(* Logix 5000 project; controller CIP_14485201 vendor 1 type 14 code 216 rev 38.11; software revision 38.01; part 5 of 12 *)
(* tags used below, declared in another part *)
   Alarm_Ack : INT[8];   // ALARMS ACKNOWLEDGE BITS
   Alarm_Present : INT[8];   // ALARM MSGS 1-127 PRESENT BITS
   Alarm_Timer : TIMER[128];   // ALARM MSGS 1-127 DELAY TIMERS
(* MainProgram, continued *)

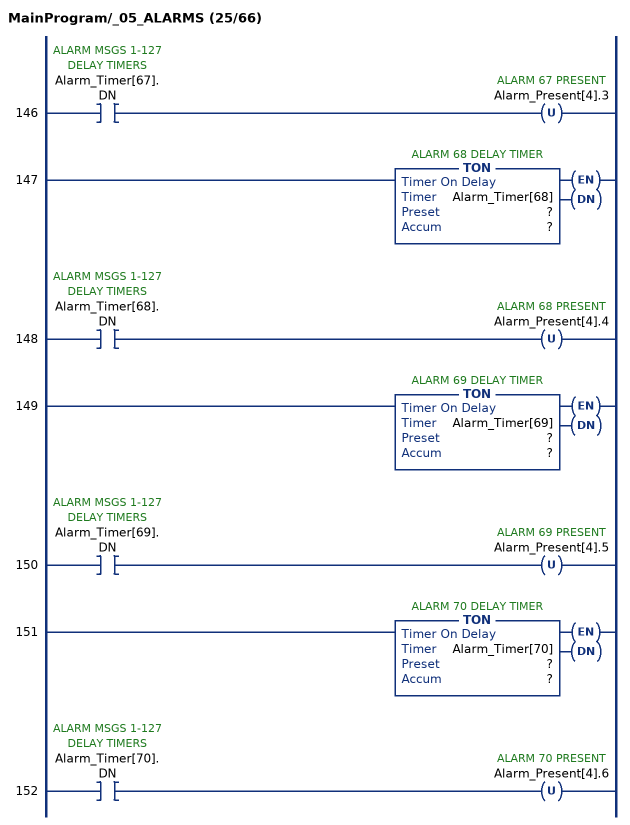
   [picture p52: MainProgram/_05_ALARMS rungs 146-152]
   146: XIC(Alarm_Timer[67].DN)OTU(Alarm_Present[4].3);
   147: TON(Alarm_Timer[68],?,?);
   148: XIC(Alarm_Timer[68].DN)OTU(Alarm_Present[4].4);
   149: TON(Alarm_Timer[69],?,?);
   150: XIC(Alarm_Timer[69].DN)OTU(Alarm_Present[4].5);
   151: TON(Alarm_Timer[70],?,?);
   152: XIC(Alarm_Timer[70].DN)OTU(Alarm_Present[4].6);
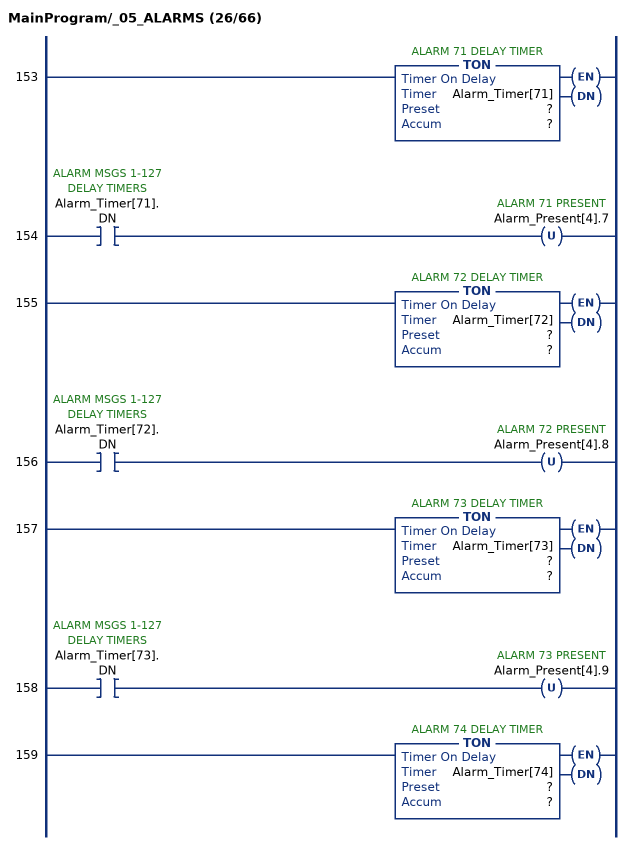
   153: TON(Alarm_Timer[71],?,?);
   154: XIC(Alarm_Timer[71].DN)OTU(Alarm_Present[4].7);
   155: TON(Alarm_Timer[72],?,?);
   156: XIC(Alarm_Timer[72].DN)OTU(Alarm_Present[4].8);
   157: TON(Alarm_Timer[73],?,?);
   158: XIC(Alarm_Timer[73].DN)OTU(Alarm_Present[4].9);
   159: TON(Alarm_Timer[74],?,?);
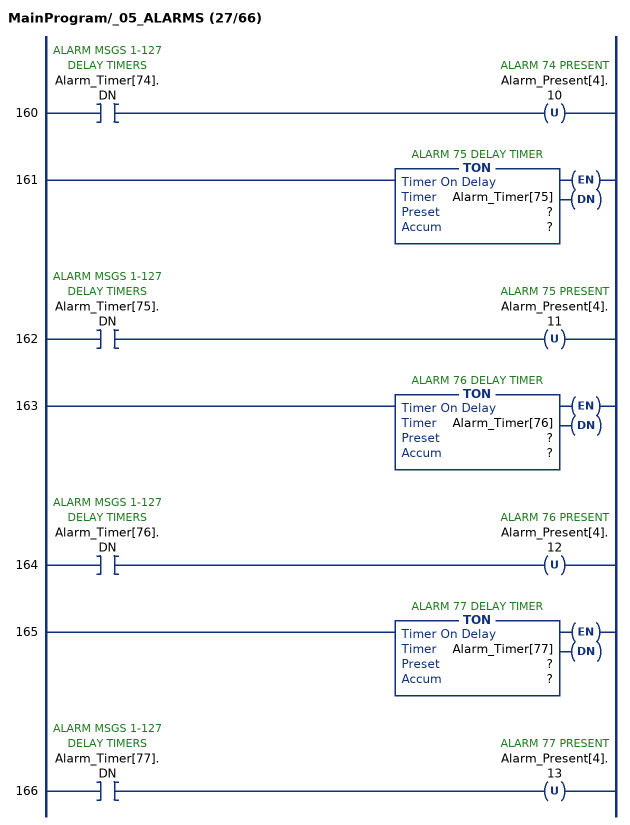
   160: XIC(Alarm_Timer[74].DN)OTU(Alarm_Present[4].10);
   161: TON(Alarm_Timer[75],?,?);
   162: XIC(Alarm_Timer[75].DN)OTU(Alarm_Present[4].11);
   163: TON(Alarm_Timer[76],?,?);
   164: XIC(Alarm_Timer[76].DN)OTU(Alarm_Present[4].12);
   165: TON(Alarm_Timer[77],?,?);
   166: XIC(Alarm_Timer[77].DN)OTU(Alarm_Present[4].13);
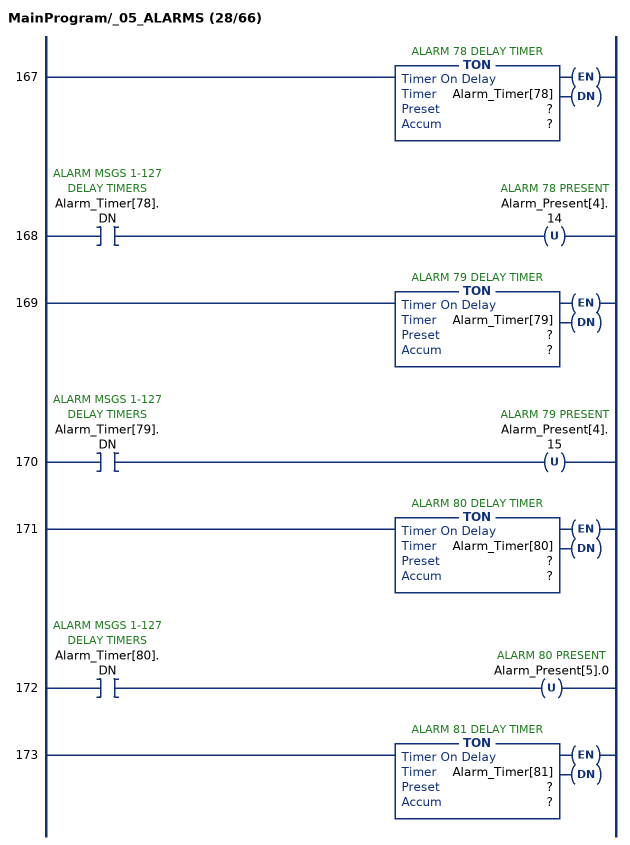
   167: TON(Alarm_Timer[78],?,?);
   168: XIC(Alarm_Timer[78].DN)OTU(Alarm_Present[4].14);
   169: TON(Alarm_Timer[79],?,?);
   170: XIC(Alarm_Timer[79].DN)OTU(Alarm_Present[4].15);
   171: TON(Alarm_Timer[80],?,?);
   172: XIC(Alarm_Timer[80].DN)OTU(Alarm_Present[5].0);
   173: TON(Alarm_Timer[81],?,?);
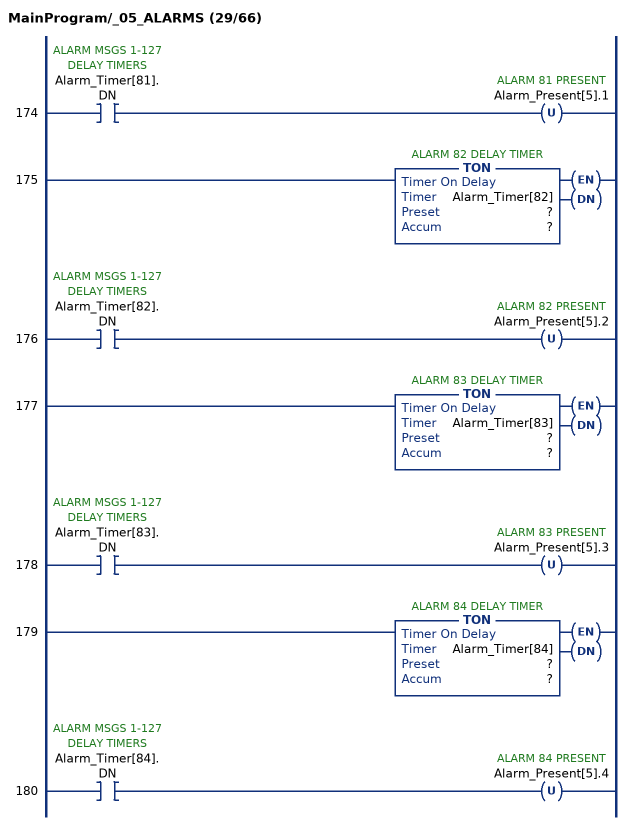
   174: XIC(Alarm_Timer[81].DN)OTU(Alarm_Present[5].1);
   175: TON(Alarm_Timer[82],?,?);
   176: XIC(Alarm_Timer[82].DN)OTU(Alarm_Present[5].2);
   177: TON(Alarm_Timer[83],?,?);
   178: XIC(Alarm_Timer[83].DN)OTU(Alarm_Present[5].3);
   179: TON(Alarm_Timer[84],?,?);
   180: XIC(Alarm_Timer[84].DN)OTU(Alarm_Present[5].4);
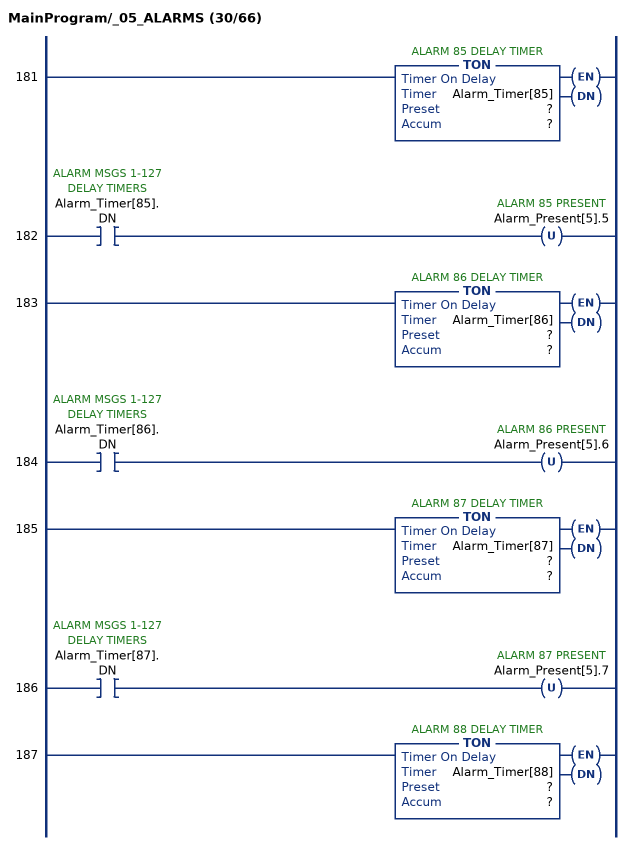
   181: TON(Alarm_Timer[85],?,?);
   182: XIC(Alarm_Timer[85].DN)OTU(Alarm_Present[5].5);
   183: TON(Alarm_Timer[86],?,?);
   184: XIC(Alarm_Timer[86].DN)OTU(Alarm_Present[5].6);
   185: TON(Alarm_Timer[87],?,?);
   186: XIC(Alarm_Timer[87].DN)OTU(Alarm_Present[5].7);
   187: TON(Alarm_Timer[88],?,?);
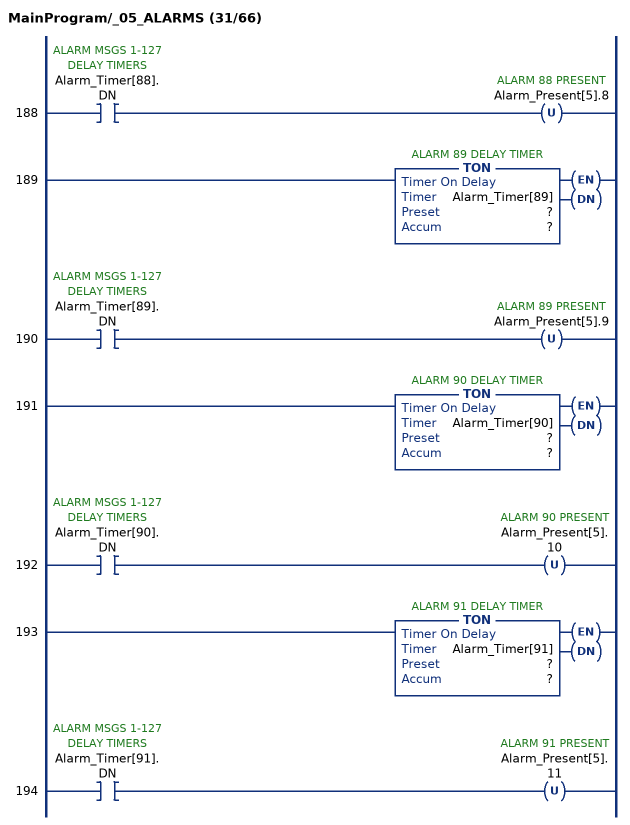
   188: XIC(Alarm_Timer[88].DN)OTU(Alarm_Present[5].8);
   189: TON(Alarm_Timer[89],?,?);
   190: XIC(Alarm_Timer[89].DN)OTU(Alarm_Present[5].9);
   191: TON(Alarm_Timer[90],?,?);
   192: XIC(Alarm_Timer[90].DN)OTU(Alarm_Present[5].10);
   193: TON(Alarm_Timer[91],?,?);
   194: XIC(Alarm_Timer[91].DN)OTU(Alarm_Present[5].11);
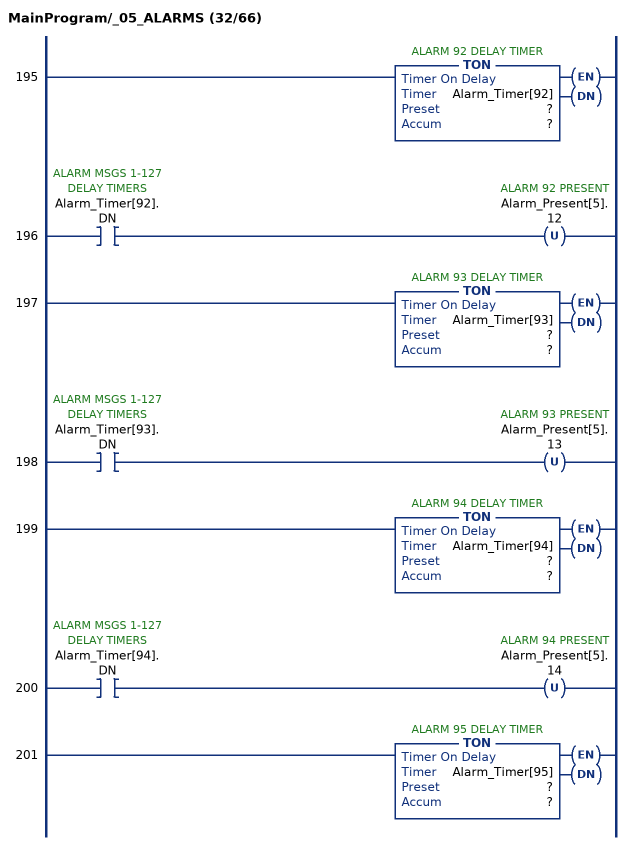
   195: TON(Alarm_Timer[92],?,?);
   196: XIC(Alarm_Timer[92].DN)OTU(Alarm_Present[5].12);
   197: TON(Alarm_Timer[93],?,?);
   198: XIC(Alarm_Timer[93].DN)OTU(Alarm_Present[5].13);
   199: TON(Alarm_Timer[94],?,?);
   200: XIC(Alarm_Timer[94].DN)OTU(Alarm_Present[5].14);
   201: TON(Alarm_Timer[95],?,?);
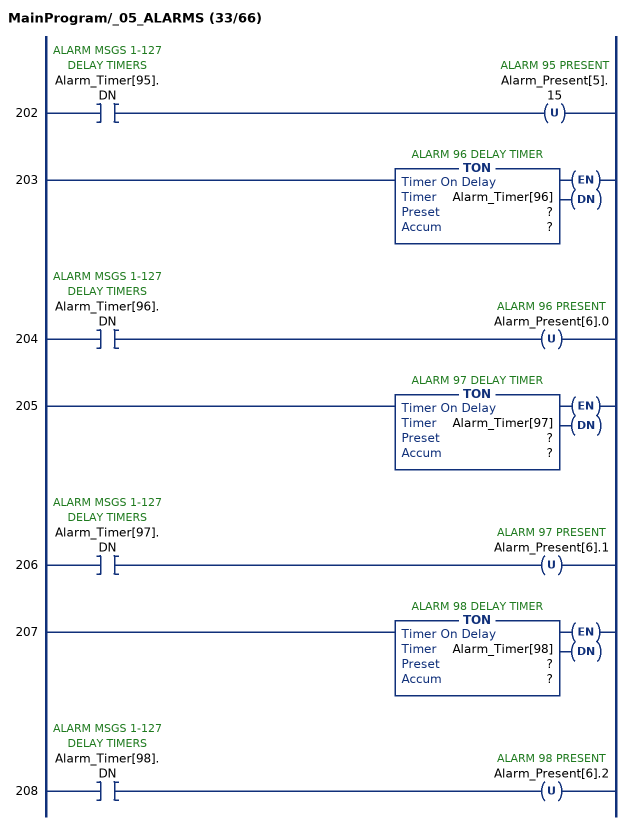
   202: XIC(Alarm_Timer[95].DN)OTU(Alarm_Present[5].15);
   203: TON(Alarm_Timer[96],?,?);
   204: XIC(Alarm_Timer[96].DN)OTU(Alarm_Present[6].0);
   205: TON(Alarm_Timer[97],?,?);
   206: XIC(Alarm_Timer[97].DN)OTU(Alarm_Present[6].1);
   207: TON(Alarm_Timer[98],?,?);
   208: XIC(Alarm_Timer[98].DN)OTU(Alarm_Present[6].2);
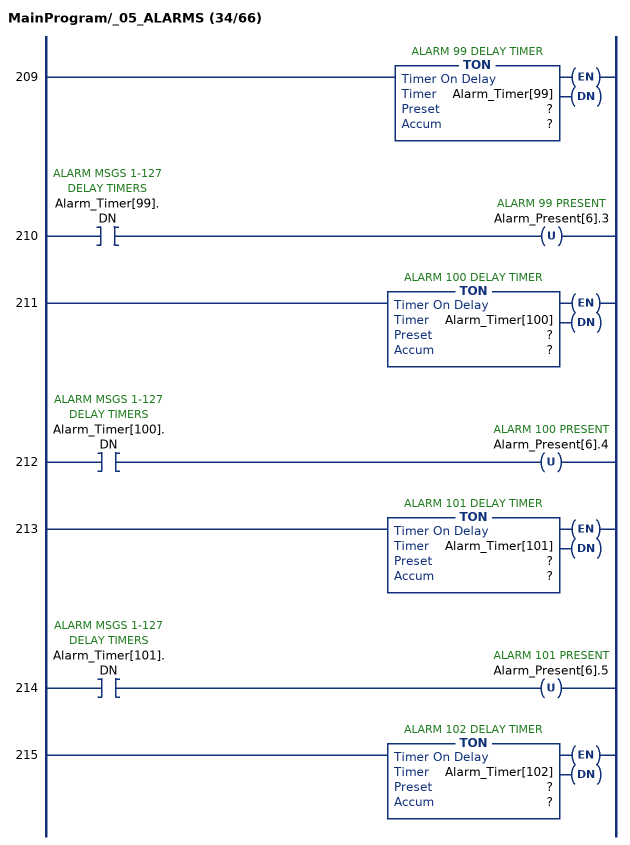
   209: TON(Alarm_Timer[99],?,?);
   210: XIC(Alarm_Timer[99].DN)OTU(Alarm_Present[6].3);
   211: TON(Alarm_Timer[100],?,?);
   212: XIC(Alarm_Timer[100].DN)OTU(Alarm_Present[6].4);
   213: TON(Alarm_Timer[101],?,?);
   214: XIC(Alarm_Timer[101].DN)OTU(Alarm_Present[6].5);
   215: TON(Alarm_Timer[102],?,?);
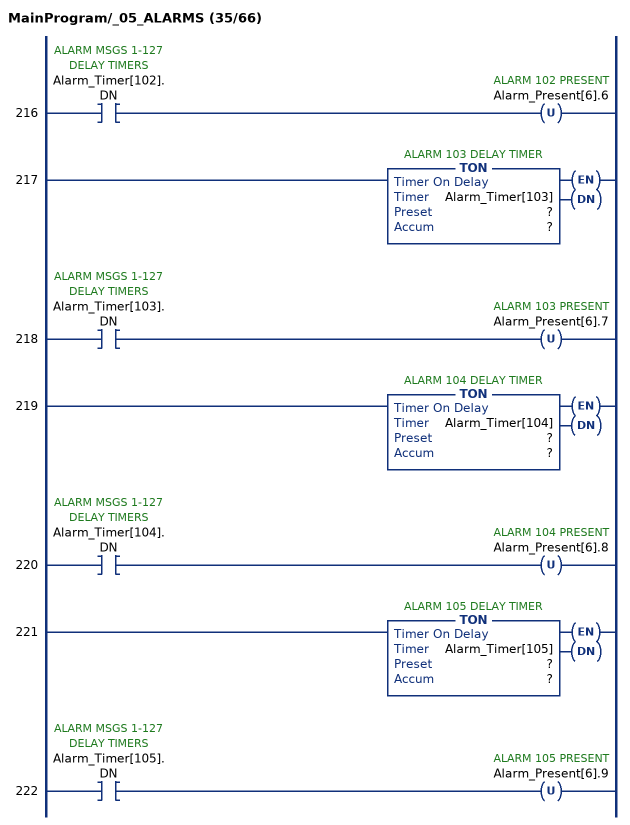
   216: XIC(Alarm_Timer[102].DN)OTU(Alarm_Present[6].6);
   217: TON(Alarm_Timer[103],?,?);
   218: XIC(Alarm_Timer[103].DN)OTU(Alarm_Present[6].7);
   219: TON(Alarm_Timer[104],?,?);
   220: XIC(Alarm_Timer[104].DN)OTU(Alarm_Present[6].8);
   221: TON(Alarm_Timer[105],?,?);
   222: XIC(Alarm_Timer[105].DN)OTU(Alarm_Present[6].9);
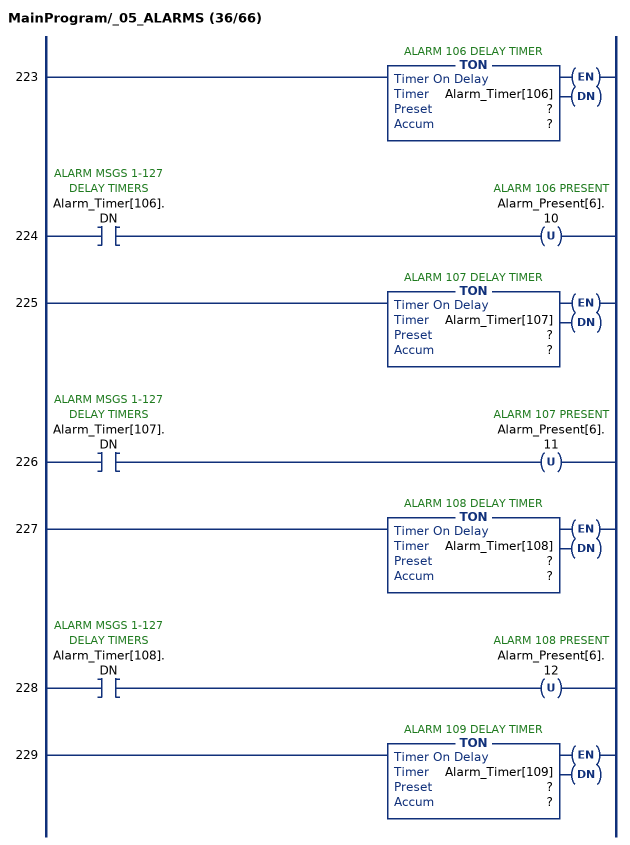
   223: TON(Alarm_Timer[106],?,?);
   224: XIC(Alarm_Timer[106].DN)OTU(Alarm_Present[6].10);
   225: TON(Alarm_Timer[107],?,?);
   226: XIC(Alarm_Timer[107].DN)OTU(Alarm_Present[6].11);
   227: TON(Alarm_Timer[108],?,?);
   228: XIC(Alarm_Timer[108].DN)OTU(Alarm_Present[6].12);
   229: TON(Alarm_Timer[109],?,?);
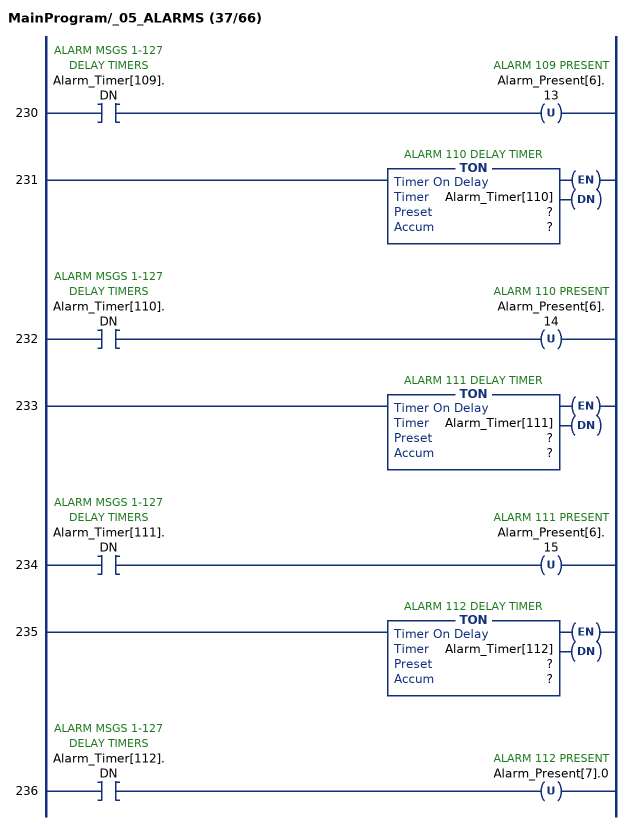
   230: XIC(Alarm_Timer[109].DN)OTU(Alarm_Present[6].13);
   231: TON(Alarm_Timer[110],?,?);
   232: XIC(Alarm_Timer[110].DN)OTU(Alarm_Present[6].14);
   233: TON(Alarm_Timer[111],?,?);
   234: XIC(Alarm_Timer[111].DN)OTU(Alarm_Present[6].15);
   235: TON(Alarm_Timer[112],?,?);
   236: XIC(Alarm_Timer[112].DN)OTU(Alarm_Present[7].0);
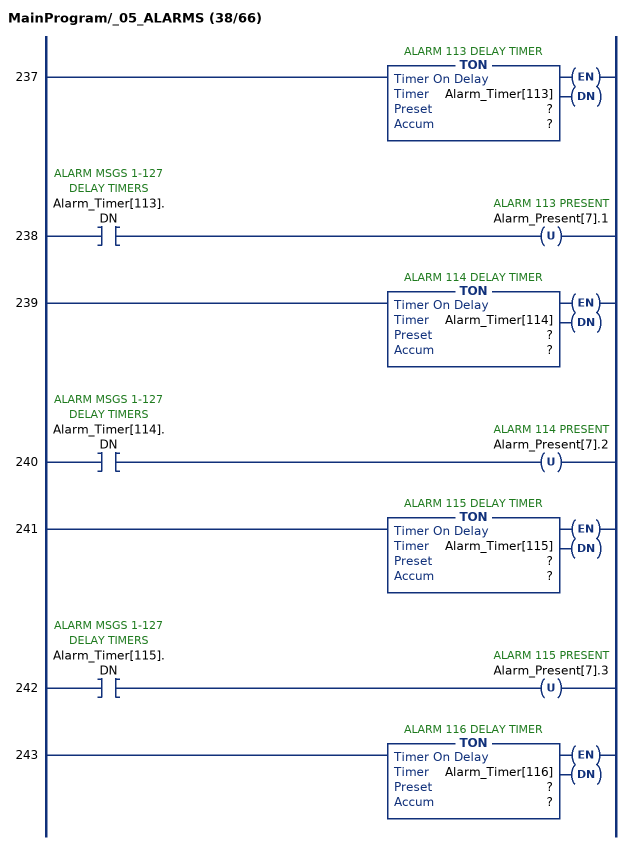
   237: TON(Alarm_Timer[113],?,?);
   238: XIC(Alarm_Timer[113].DN)OTU(Alarm_Present[7].1);
   239: TON(Alarm_Timer[114],?,?);
   240: XIC(Alarm_Timer[114].DN)OTU(Alarm_Present[7].2);
   241: TON(Alarm_Timer[115],?,?);
   242: XIC(Alarm_Timer[115].DN)OTU(Alarm_Present[7].3);
   243: TON(Alarm_Timer[116],?,?);
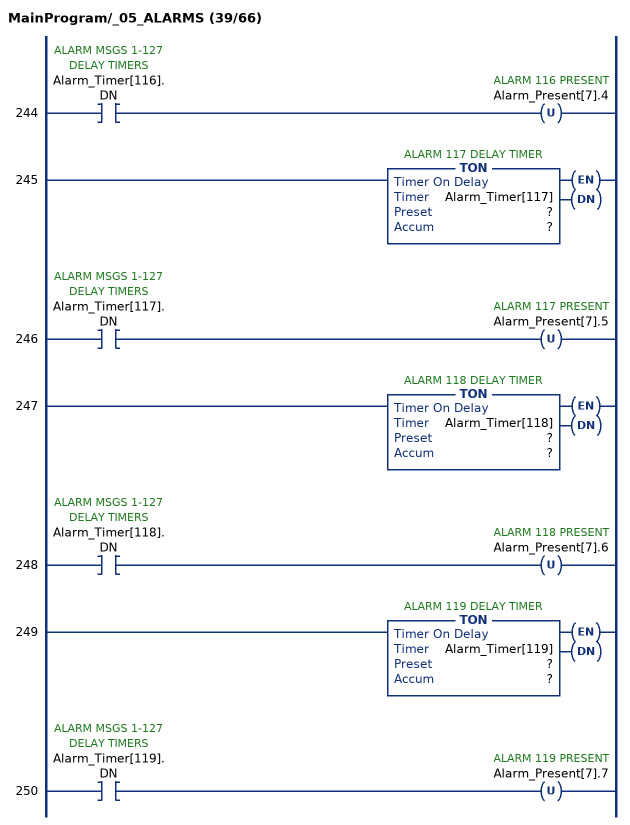
   244: XIC(Alarm_Timer[116].DN)OTU(Alarm_Present[7].4);
   245: TON(Alarm_Timer[117],?,?);
   246: XIC(Alarm_Timer[117].DN)OTU(Alarm_Present[7].5);
   247: TON(Alarm_Timer[118],?,?);
   248: XIC(Alarm_Timer[118].DN)OTU(Alarm_Present[7].6);
   249: TON(Alarm_Timer[119],?,?);
   250: XIC(Alarm_Timer[119].DN)OTU(Alarm_Present[7].7);
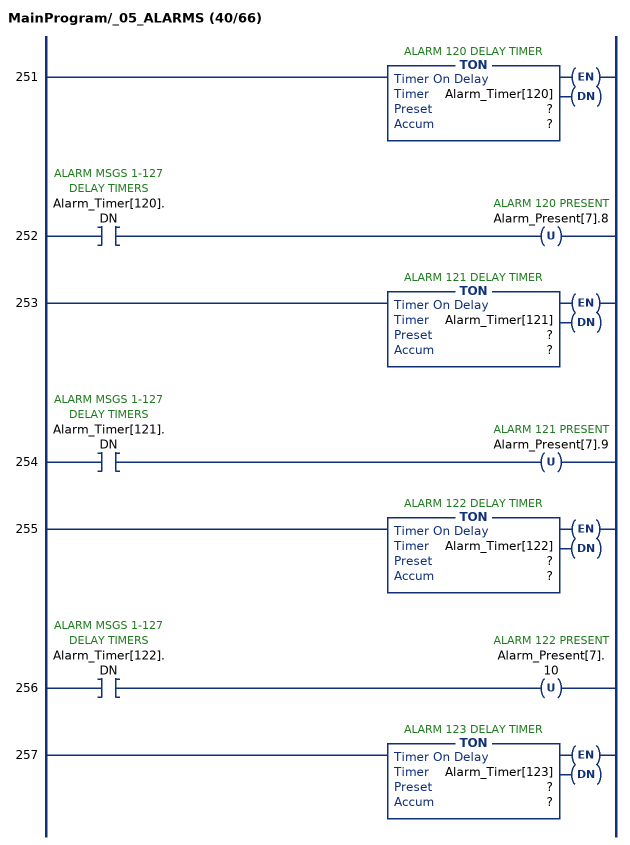
   251: TON(Alarm_Timer[120],?,?);
   252: XIC(Alarm_Timer[120].DN)OTU(Alarm_Present[7].8);
   253: TON(Alarm_Timer[121],?,?);
   254: XIC(Alarm_Timer[121].DN)OTU(Alarm_Present[7].9);
   255: TON(Alarm_Timer[122],?,?);
   256: XIC(Alarm_Timer[122].DN)OTU(Alarm_Present[7].10);
   257: TON(Alarm_Timer[123],?,?);
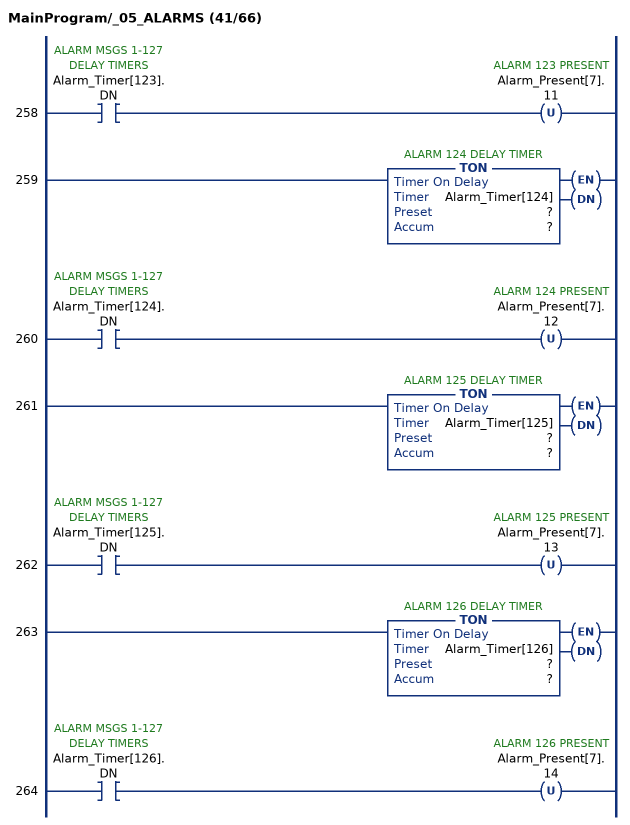
   258: XIC(Alarm_Timer[123].DN)OTU(Alarm_Present[7].11);
   259: TON(Alarm_Timer[124],?,?);
   260: XIC(Alarm_Timer[124].DN)OTU(Alarm_Present[7].12);
   261: TON(Alarm_Timer[125],?,?);
   262: XIC(Alarm_Timer[125].DN)OTU(Alarm_Present[7].13);
   263: TON(Alarm_Timer[126],?,?);
   264: XIC(Alarm_Timer[126].DN)OTU(Alarm_Present[7].14);
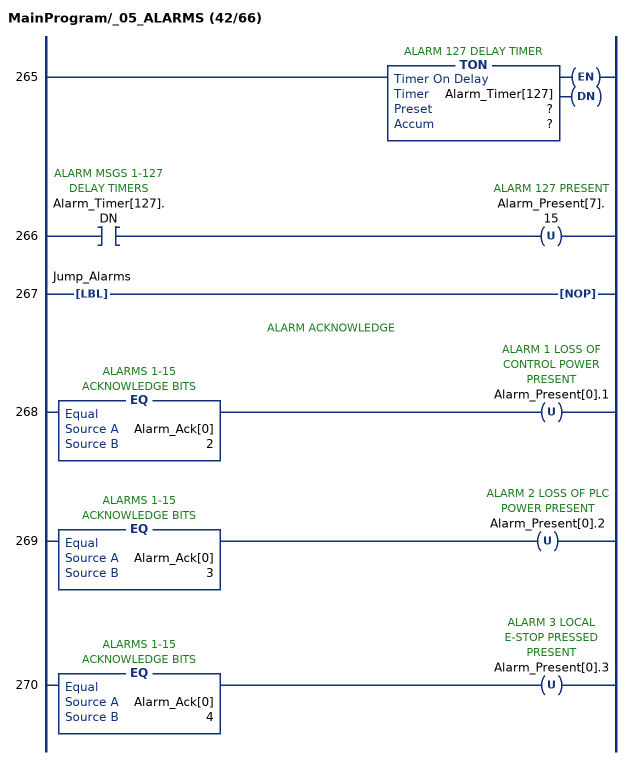
   265: TON(Alarm_Timer[127],?,?);
   266: XIC(Alarm_Timer[127].DN)OTU(Alarm_Present[7].15);
   267: LBL(Jump_Alarms)NOP();
   // ALARM ACKNOWLEDGE
   268: EQ(Alarm_Ack[0],2)OTU(Alarm_Present[0].1);
   269: EQ(Alarm_Ack[0],3)OTU(Alarm_Present[0].2);
   270: EQ(Alarm_Ack[0],4)OTU(Alarm_Present[0].3);
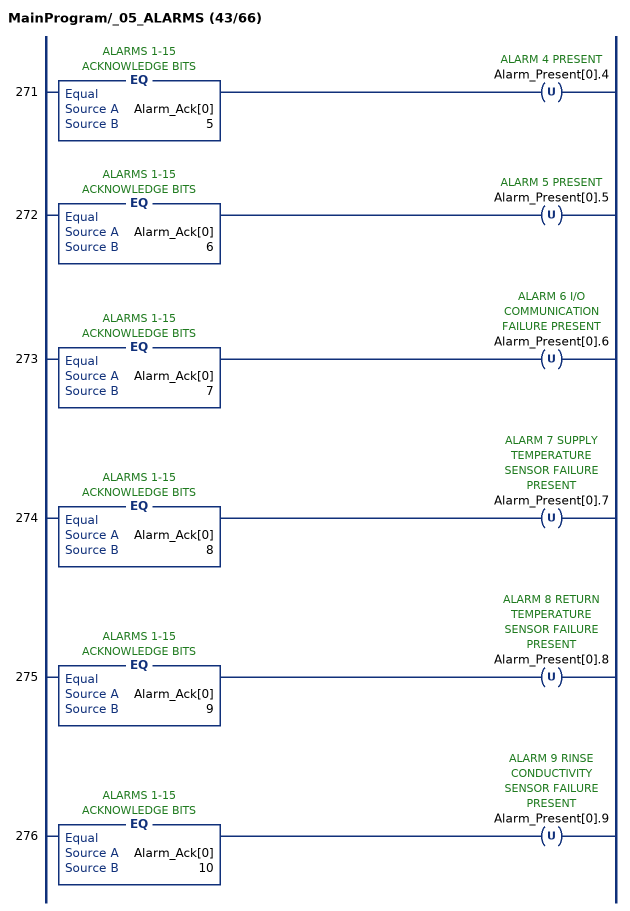
   271: EQ(Alarm_Ack[0],5)OTU(Alarm_Present[0].4);
   272: EQ(Alarm_Ack[0],6)OTU(Alarm_Present[0].5);
   273: EQ(Alarm_Ack[0],7)OTU(Alarm_Present[0].6);
   274: EQ(Alarm_Ack[0],8)OTU(Alarm_Present[0].7);
   275: EQ(Alarm_Ack[0],9)OTU(Alarm_Present[0].8);
   276: EQ(Alarm_Ack[0],10)OTU(Alarm_Present[0].9);
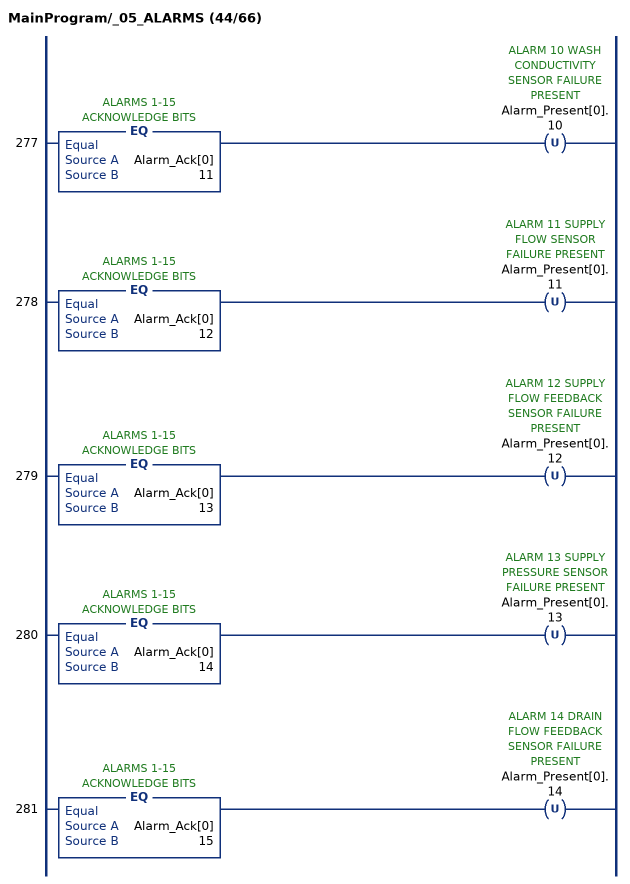
   277: EQ(Alarm_Ack[0],11)OTU(Alarm_Present[0].10);
   278: EQ(Alarm_Ack[0],12)OTU(Alarm_Present[0].11);
   279: EQ(Alarm_Ack[0],13)OTU(Alarm_Present[0].12);
   280: EQ(Alarm_Ack[0],14)OTU(Alarm_Present[0].13);
   281: EQ(Alarm_Ack[0],15)OTU(Alarm_Present[0].14);
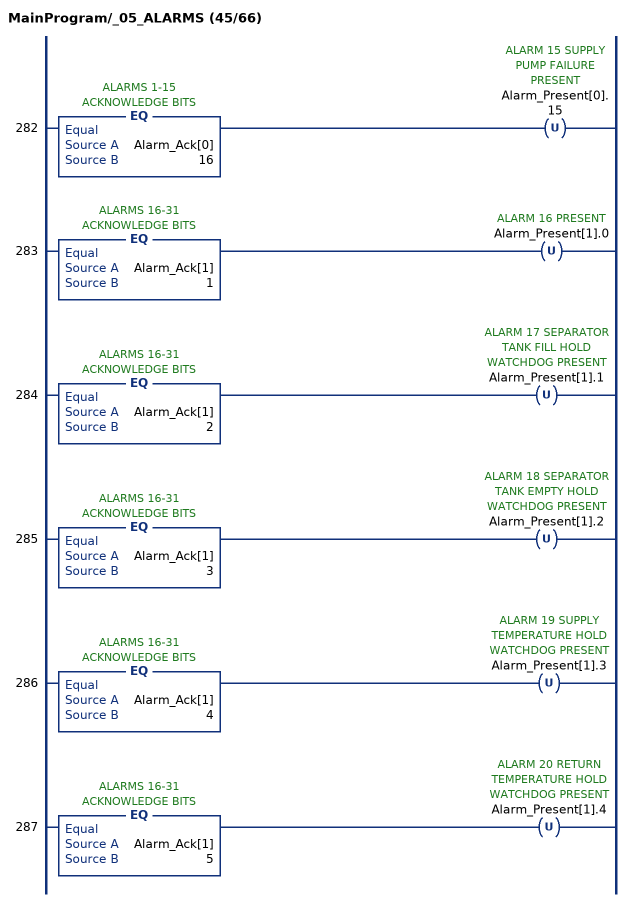
   282: EQ(Alarm_Ack[0],16)OTU(Alarm_Present[0].15);
   283: EQ(Alarm_Ack[1],1)OTU(Alarm_Present[1].0);
   284: EQ(Alarm_Ack[1],2)OTU(Alarm_Present[1].1);
   285: EQ(Alarm_Ack[1],3)OTU(Alarm_Present[1].2);
   286: EQ(Alarm_Ack[1],4)OTU(Alarm_Present[1].3);
   287: EQ(Alarm_Ack[1],5)OTU(Alarm_Present[1].4);
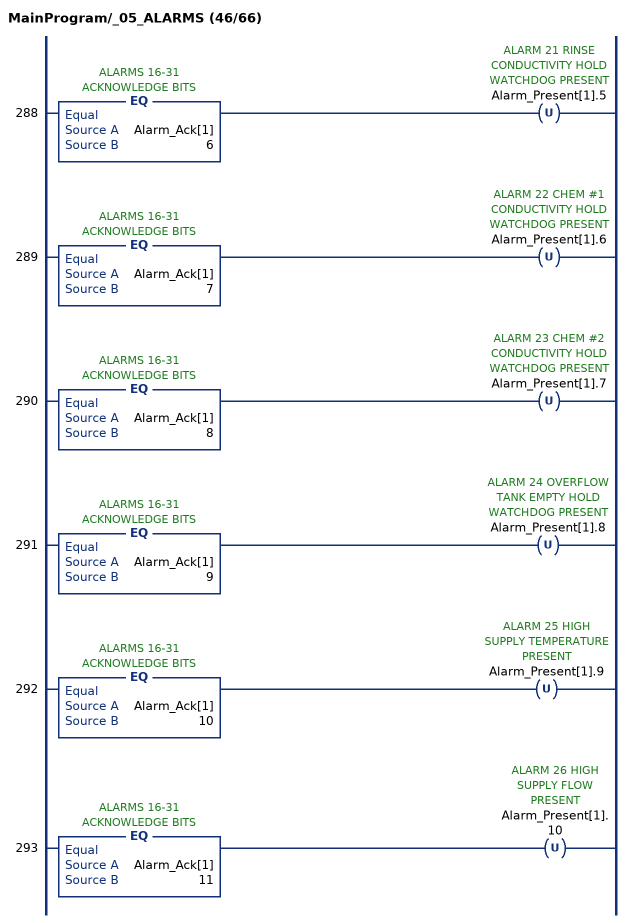
   288: EQ(Alarm_Ack[1],6)OTU(Alarm_Present[1].5);
   289: EQ(Alarm_Ack[1],7)OTU(Alarm_Present[1].6);
   290: EQ(Alarm_Ack[1],8)OTU(Alarm_Present[1].7);
   291: EQ(Alarm_Ack[1],9)OTU(Alarm_Present[1].8);
   292: EQ(Alarm_Ack[1],10)OTU(Alarm_Present[1].9);
   293: EQ(Alarm_Ack[1],11)OTU(Alarm_Present[1].10);
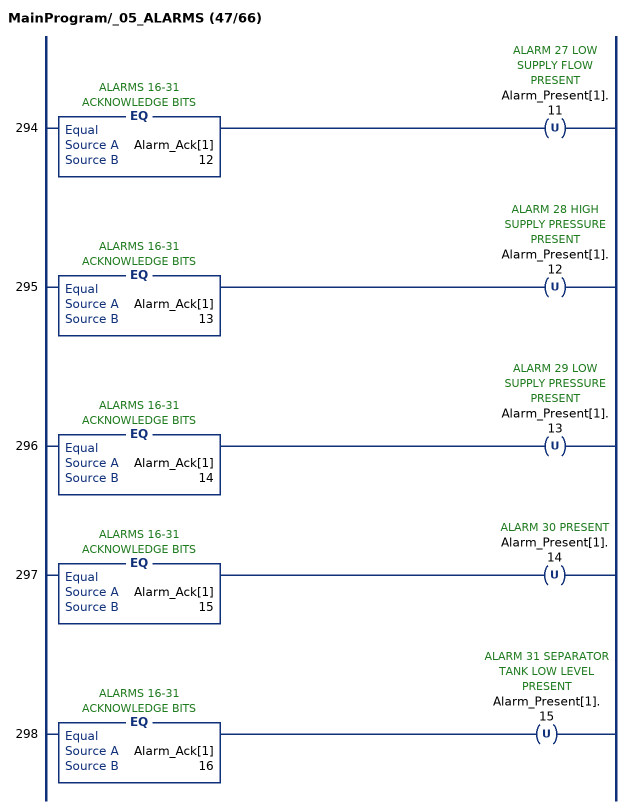
   294: EQ(Alarm_Ack[1],12)OTU(Alarm_Present[1].11);
   295: EQ(Alarm_Ack[1],13)OTU(Alarm_Present[1].12);
   296: EQ(Alarm_Ack[1],14)OTU(Alarm_Present[1].13);
   297: EQ(Alarm_Ack[1],15)OTU(Alarm_Present[1].14);
   298: EQ(Alarm_Ack[1],16)OTU(Alarm_Present[1].15);
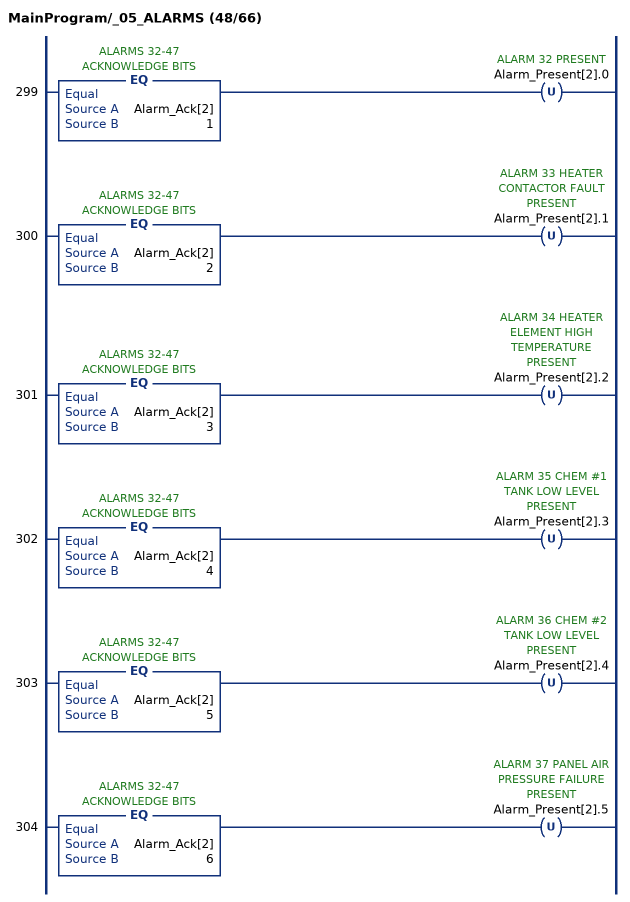
   299: EQ(Alarm_Ack[2],1)OTU(Alarm_Present[2].0);
   300: EQ(Alarm_Ack[2],2)OTU(Alarm_Present[2].1);
   301: EQ(Alarm_Ack[2],3)OTU(Alarm_Present[2].2);
   302: EQ(Alarm_Ack[2],4)OTU(Alarm_Present[2].3);
   303: EQ(Alarm_Ack[2],5)OTU(Alarm_Present[2].4);
   304: EQ(Alarm_Ack[2],6)OTU(Alarm_Present[2].5);
